// TIA Portal V20 export
DATA_BLOCK "HMI_Signale"   // DB500
{ S7_Optimized_Access := 'FALSE' }
// stored: AutoNumber false
   VAR RETAIN
      Statistik_BA : Bool := FALSE;   // Anforderung kommt von HMI
      Automatik_BA : Bool := FALSE;   // Anforderung kommt von HMI
      Manuell_BA : Bool := FALSE;   // Anforderung kommt von HMI
      Verwalten_BA : Bool := FALSE;   // Anforderung kommt von HMI
      Richten_BA : Bool := FALSE;   // Anforderung kommt von HMI
      Dauer_Manuell_Betrieb : Bool := TRUE;   // Dauerbetrieb = 1 / Manuellbetrieb = 0
      Stop_nach_Zyklus : Bool := FALSE;
      Ablauf_aktiv : Bool := FALSE;
      Leerfahren_angewaehlt : Bool := FALSE;
      Leerfahren_Laeuft : Bool := FALSE;
      Leerfahren_ende : Bool := FALSE;
      Freigabe_Zyklus : Bool := FALSE;   // Zyklus Freigegeben
      FPStarttaste : Bool := FALSE;
      Stop_Von_Stoermeldung : Bool := FALSE;
      Sammelstoerung : Bool := FALSE;
      SK_aktiv : Bool;   // min 1 Schrittkettenablauf ist aktiv
   END_VAR
BEGIN
END_DATA_BLOCK
